(* IEC 61131-3 sources: ieccompiler/test/syn_tests, 17 files *)

(* ---- test_func.st ---- *)
FUNCTION test_func
  VAR
    b_Start_Stop : DINT;
    N : DINT;
  END_VAR

  IF b_Start_Stop > 0 THEN
    N := N + 7;
  ELSIF b_Start_Stop > 111111 AND N < 222222 AND (N > 333333 AND N < 444444) AND N <> 555555 THEN
    N := N + 8;
  ELSE
    N := N + 9;
  END_IF
END_FUNCTION

(* ---- test_fb.st ---- *)
FUNCTION_BLOCK test_fb
  VAR
    b_Start_Stop:DINT;
    N : DINT := 10;
  END_VAR

  IF b_Start_Stop > 0 THEN
    N := N + 7;
  ELSIF b_Start_Stop > 111111
    AND N < 222222
    AND (N > 333333 AND N < 444444)
    AND N <> 555555 THEN
    N := N + 8;
  ELSE
    N := N + 9;
  END_IF
END_FUNCTION_BLOCK

(* ---- main.st ---- *)
IMPORT test_if.st
IMPORT test_and.st
IMPORT test_or.st
IMPORT test_while.st
IMPORT test_fb.st
IMPORT test_func.st
IMPORT test_arithmetic.st
IMPORT test_paren.st
IMPORT test_parenno.st
IMPORT test_paren_nest.st
IMPORT test_priority.st
IMPORT test_typecheck.st
IMPORT test_xor.st
//IMPORT test_func_return.st
//IMPORT test_not.st
//IMPORT test_func_for.st
IMPORT test_repeat.st
//IMPORT test_case.st
//IMPORT test_compare.st
PROGRAM main
END_PROGRAM

(* ---- test_and.st ---- *)
PROGRAM test_and
  VAR
    b_Start_Stop : DINT;
    N : DINT;
  END_VAR

  IF b_Start_Stop > 111111 AND N < 222222 THEN
    N := N + 7;
  ELSIF b_Start_Stop > 111111 THEN
    N := N + 8;
  ELSE
    N := N + 9;
  END_IF
END_PROGRAM

(* ---- test_arithmetic.st ---- *)
PROGRAM test_arithmetic
  VAR
    A : INT;
    B : INT;
    C : INT;
  END_VAR

  C := A + B - 9;
  C := A - B + 9;
  C := A * B / 2;
  C := A / 2 * B;
  C := B + 5 - 2 * B / C;
END_PROGRAM

(* ---- test_func_return.st ---- *)
PROGRAM test_func_return
  VAR
    B : INT;
    C : INT;
    D : BOOL;
  END_VAR

  D := test_func_return_add(B,C);
END_PROGRAM

FUNCTION test_func_return_add : INT
  VAR
    KK : INT;
    VV : BOOL;
  END_VAR

  VAR_INPUT
    BBB : INT;
    CCC : INT;
  END_VAR

  KK := BBB + CCC + 9;
  RETURN KK;
END_FUNCTION

(* ---- test_if.st ---- *)
PROGRAM test_if
  VAR
    b_Start_Stop : DINT;
    N : DINT;
  END_VAR

  IF b_Start_Stop > 0 THEN
    N := N + 7;
  ELSIF b_Start_Stop > 111111 THEN
    N := N + 8;
  ELSE
    N := N + 9;
  END_IF
END_PROGRAM

(* ---- test_not.st ---- *)
PROGRAM test_not
  VAR
    b_Start_Stop : DINT;
    N : DINT;
    bFlag : BOOL;
  END_VAR

  IF NOT bFlag THEN
    N := N + 7;
  ELSE
    N := N + 9;
  END_IF
END_PROGRAM

(* ---- test_or.st ---- *)
PROGRAM test_or
  VAR
    b_Start_Stop : DINT;
    N : DINT;
  END_VAR

  IF b_Start_Stop > 111111 OR N < 222222 THEN
    N := N + 7;
  ELSIF b_Start_Stop > 333333 THEN
    N := N + 8;
  ELSE
    N := N + 9;
  END_IF
END_PROGRAM

(* ---- test_paren.st ---- *)
PROGRAM test_paren
  VAR
    b_Start_Stop : DINT;
    N : DINT;
  END_VAR

  IF b_Start_Stop > 111111 AND ( b_Start_Stop < 222222 OR  b_Start_Stop < 333000) THEN
    N := N + 7;
  ELSIF b_Start_Stop > 333333 OR ( b_Start_Stop < 111111 AND  b_Start_Stop > 5) THEN
    N := N + 8;
  ELSE
    N := N + 9;
  END_IF
END_PROGRAM

(* ---- test_paren_nest.st ---- *)
PROGRAM test_paren_nest
  VAR
    A : INT;
  END_VAR
  A := A*(A/(A+ 2)+3);
  A := A*(A/(A+2) );//ok
  A := A*(A/(A+2));//Invalid syntax
  A := A*( (A+2)*3);//ok
  A := A*((A+2)*3);//Invalid syntax
END_PROGRAM

(* ---- test_parenno.st ---- *)
PROGRAM test_parenno
  VAR
    b_Start_Stop: DINT;
    N: DINT;
  END_VAR

  IF b_Start_Stop > 111111 AND  b_Start_Stop < 222222 OR  b_Start_Stop < 333000 THEN
    N := N + 7;
  ELSIF b_Start_Stop > 333333 OR b_Start_Stop < 111111 AND  b_Start_Stop > 5 THEN
    N := N + 8;
  ELSE
    N := N + 9;
  END_IF
END_PROGRAM

(* ---- test_priority.st ---- *)
PROGRAM test_priority
  VAR
    b_Start_Stop: DINT;
    N: DINT;
  END_VAR

  WHILE b_Start_Stop  > 200 OR b_Start_Stop < 111111 AND N < 222222 DO
    N := N + 10;
    N := b_Start_Stop+5-2*b_Start_Stop/N;
  END_WHILE
END_PROGRAM

(* ---- test_repeat.st ---- *)
PROGRAM test_repeat
  VAR
    i  : INT;
  END_VAR

  REPEAT
    i := i + 1;
  UNTIL i = 4;
  END_REPEAT
END_PROGRAM

(* ---- test_typecheck.st ---- *)
PROGRAM test_typecheckend_type
  VAR
    B: INT;
    C: INT;
    D: BOOL;
  END_VAR

  C := functest(D, B);
END_PROGRAM

FUNCTION functest:INT
  VAR
    KK: INT;
  END_VAR
  VAR_INPUT
    bFlag: BOOL;
    nIndex: INT;
  END_VAR

  IF bFlag <> 0 THEN
    KK := nIndex + 1;
  END_IF
END_FUNCTION

(* ---- test_while.st ---- *)
PROGRAM test_while
  VAR
    b_Start_Stop: DINT;
    N: DINT;
  END_VAR

  WHILE b_Start_Stop  > 200 AND b_Start_Stop < 111111 OR N < 222222 DO
    N := N + 10;
  END_WHILE
END_PROGRAM

(* ---- test_xor.st ---- *)
PROGRAM test_xor
  VAR
    b_Start_Stop: DINT;
    N: DINT;
  END_VAR

  IF b_Start_Stop > 111111 XOR N < 222222 THEN
    N := N + 7;
  ELSIF b_Start_Stop > 333333 THEN
    N := N + 8;
  ELSE
    N := N + 9;
  END_IF
END_PROGRAM
